(* IEC 61131-3 sources: SemantiST/benchmarks/defects/designed/d06_service_counter/buggy, 1 file *)

(* ---- target.st ---- *)
FUNCTION_BLOCK D06_SERVICE_COUNTER
VAR_INPUT
    Run : BOOL;
    Speed : INT;
    ResetService : BOOL;
END_VAR
VAR_OUTPUT
    Hours : INT;
    ServiceDue : BOOL;
    Interval : INT;
END_VAR
VAR
    plan : ARRAY[0..11] OF INT := [50, 50, 100, 100, 100, 200, 200, 200, 400, 400, 400, 800];
END_VAR

IF ResetService THEN
    Hours := 0;
ELSIF Run AND Speed >= 1450 AND Speed <= 1550 THEN
    Hours := Hours + 1;
END_IF;
IF Hours >= 10 THEN
    (* defect: Hours / 10 is not clamped to the 12-entry plan; Hours = 120 reads plan[12] *)
    Interval := plan[Hours / 10];
    ServiceDue := Hours MOD 10 = 0;
END_IF;
END_FUNCTION_BLOCK
